Fanuc KAREL source: kt00366.KL

-- PROVISIONAL review KL for V770-1; original PC SHA256 80827090fef683ad164372d2d90eec2788ff83400dc677b4cfa629a780ac50b8
-- Incomplete behavior may be omitted. Consult companion uncertainty JSON. Do not deploy.
PROGRAM KT00366
%NOLOCKGROUP
VAR
  I1 : INTEGER
  R2 : REAL
  OUT : BOOLEAN
BEGIN
  -- UNRESOLVED_PC offsets 5-16; opcodes 2E,23
  -- UNRESOLVED_PC offsets 21-32; opcodes 2E,23
  -- UNRESOLVED_PC offsets 37-59; opcodes 21,21,29,64,29,70,23
  -- UNRESOLVED_PC offsets 64-68; opcodes 7F
END KT00366
